Fanuc KAREL source: kt00038.KL

-- PROVISIONAL review KL for V770-1; original PC SHA256 bdc4f579f6188e87734442d92e1be38feae0e5980ab35d28ceb6725e2b9fa952
-- Incomplete behavior may be omitted. Consult companion uncertainty JSON. Do not deploy.
PROGRAM KT00038
%NOLOCKGROUP
VAR
  I1 : INTEGER
  OUT : REAL
-- UNRESOLVED_DECL Y2 type=002018
BEGIN
  -- UNRESOLVED_PC offsets 5-16; opcodes 2E,23
  -- UNRESOLVED_PC offsets 21-35; opcodes 2E,22,9D,33,B2
  -- UNRESOLVED_PC offsets 40-63; opcodes 21,22,9D,33,B1,53,64,23
  -- UNRESOLVED_PC offsets 68-72; opcodes 7F
END KT00038
